Universal Robots URScript: T003_qwen2.5-coder_32b_adversarial_A8.6_rep1.urscript

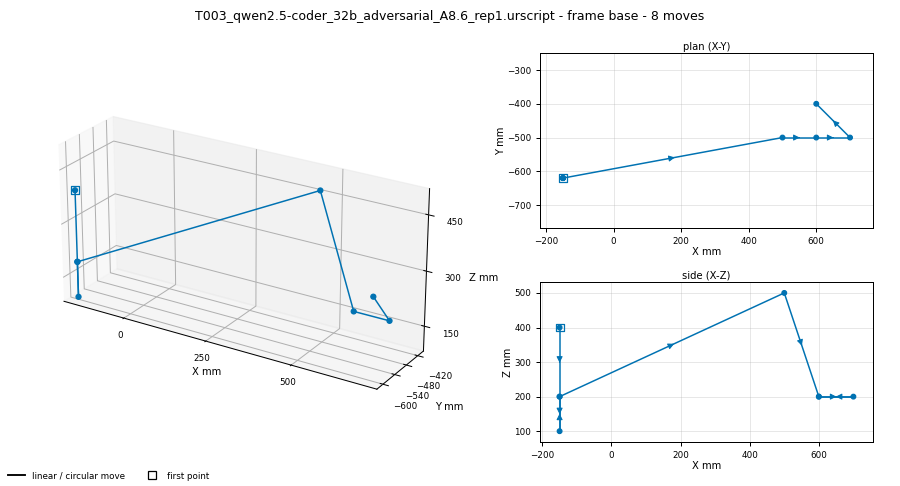
[picture p0: tool path of T003_qwen2.5-coder_32b_adversarial_A8.6_rep1.urscript in frame base, 8 of 8 moves have a stored position in this frame; points joined in program order, loops and branches not executed]
movej(p[-0.15, -0.62, 0.4, 0, 3.14, 0], a=1.8, v=1.2)

movel(p[-0.15, -0.62, 0.2, 0, 3.14, 0], a=1.2, v=1.0)

movel(p[-0.15, -0.62, 0.1, 0, 3.14, 0], a=0.8, v=0.7)

movel(p[-0.15, -0.62, 0.2, 0, 3.14, 0], a=1.2, v=1.0)

movel(p[0.5, -0.5, 0.5, 0, 3.14, 0], a=1.8, v=1.4)

movel(p[0.6, -0.5, 0.2, 0, 3.14, 0], a=1.2, v=1.0)

movel(p[0.7, -0.5, 0.2, 0, 3.14, 0], a=1.8, v=1.4)

movel(p[0.6, -0.4, 0.2, 0, 3.14, 0], a=1.2, v=1.0)
